(* Logix 5000 project; controller CIP vendor 1 type 14 code 106 rev 20.12; software revision 20.06; part 7 of 13 *)
(* tags used below, declared in another part *)
   Message_Index : ALIAS FOR Integer[30];
   Message_Present : INT[4];
   Message_SEQ : DINT[101];
   Message_Timer : TIMER[1];
   OpCode_Pin : DINT[5];
   PV_Message : DINT[3];
   SCLD_Drain_PH : REAL;
   SCLD_Dryer_Duct_Temp : REAL;
   SCLD_Dryer_Exhaust_Temp : REAL;
   SCLD_Return_Temp : REAL;
   SCLD_Rinse_Cond : REAL;
   SCLD_Solution_Tank_Lvl : REAL;
   SCLD_Solution_Tank_Lvl_Raw : REAL;
   SCLD_Supply_Flow : REAL;
   SCLD_Supply_Flow_CIP : REAL;
   SCLD_Supply_Flow_CIP100 : REAL;
   SCLD_Supply_Flow_CIP200 : REAL;
   SCLD_Supply_Pressure : REAL;
   SCLD_Supply_Temp : REAL;
   SCLD_Wash_Chamber_Lvl : REAL;
   SCLD_Wash_Chamber_Lvl_Raw : REAL;
   SCLD_Wash_Cond : REAL;
   Sequencer : CONTROL[4];
   Solution_Tank_Lvl_Calc : REAL[20];
   Solution_Tank_Lvl_Storage : REAL[3];
   Wash_Chamber_Lvl_Calc : REAL[30];
   Wash_Chamber_Lvl_Storage : REAL[3];
(* MainProgram, continued *)

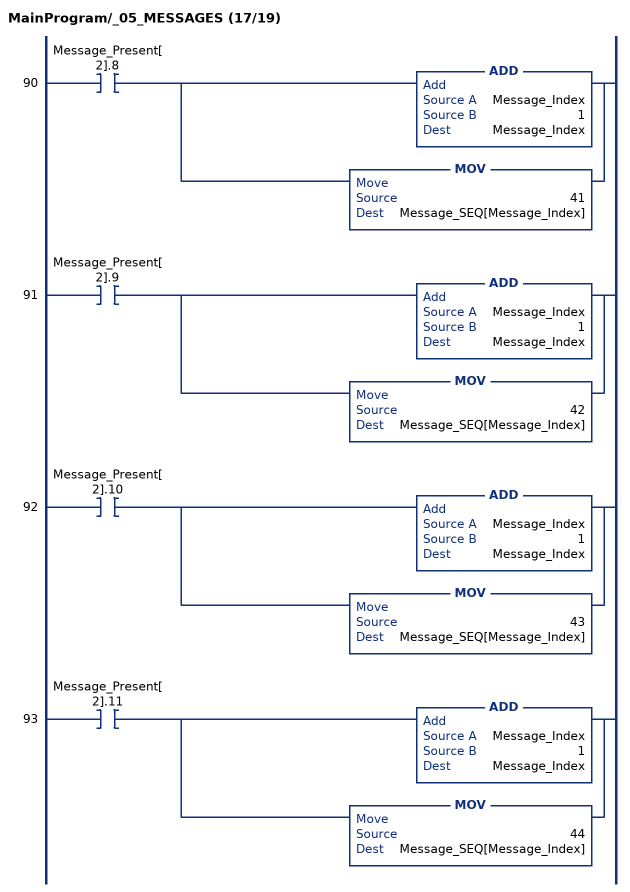
   [picture p115: MainProgram/_05_MESSAGES rungs 90-93]
   90: XIC(Message_Present[2].8)[ADD(Message_Index,1,Message_Index) ,MOV(41,Message_SEQ[Message_Index]) ];
   91: XIC(Message_Present[2].9)[ADD(Message_Index,1,Message_Index) ,MOV(42,Message_SEQ[Message_Index]) ];
   92: XIC(Message_Present[2].10)[ADD(Message_Index,1,Message_Index) ,MOV(43,Message_SEQ[Message_Index]) ];
   93: XIC(Message_Present[2].11)[ADD(Message_Index,1,Message_Index) ,MOV(44,Message_SEQ[Message_Index]) ];
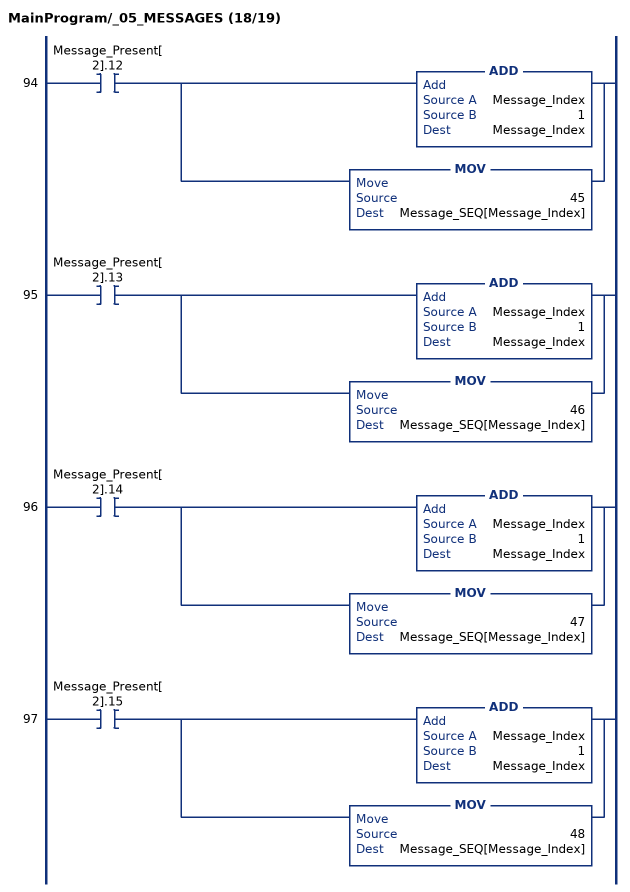
   94: XIC(Message_Present[2].12)[ADD(Message_Index,1,Message_Index) ,MOV(45,Message_SEQ[Message_Index]) ];
   95: XIC(Message_Present[2].13)[ADD(Message_Index,1,Message_Index) ,MOV(46,Message_SEQ[Message_Index]) ];
   96: XIC(Message_Present[2].14)[ADD(Message_Index,1,Message_Index) ,MOV(47,Message_SEQ[Message_Index]) ];
   97: XIC(Message_Present[2].15)[ADD(Message_Index,1,Message_Index) ,MOV(48,Message_SEQ[Message_Index]) ];
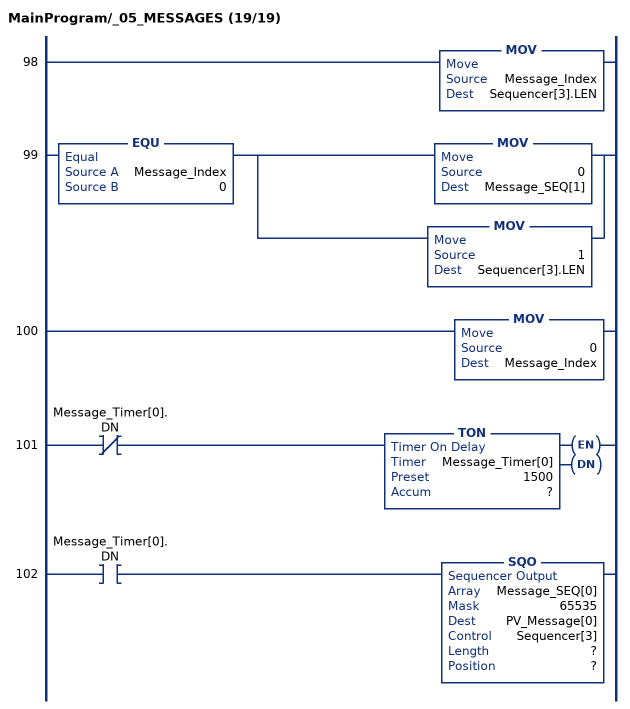
   98: MOV(Message_Index,Sequencer[3].LEN);
   99: EQU(Message_Index,0)[MOV(0,Message_SEQ[1]) ,MOV(1,Sequencer[3].LEN) ];
   100: MOV(0,Message_Index);
   101: XIO(Message_Timer[0].DN)TON(Message_Timer[0],?,?);
   102: XIC(Message_Timer[0].DN)SQO(Message_SEQ[0],65535,PV_Message[0],Sequencer[3],?,?);
END_ROUTINE

ROUTINE _07_SCALE   (* function block diagram *)
   SHEET 1   // Local Analog Input Scaling
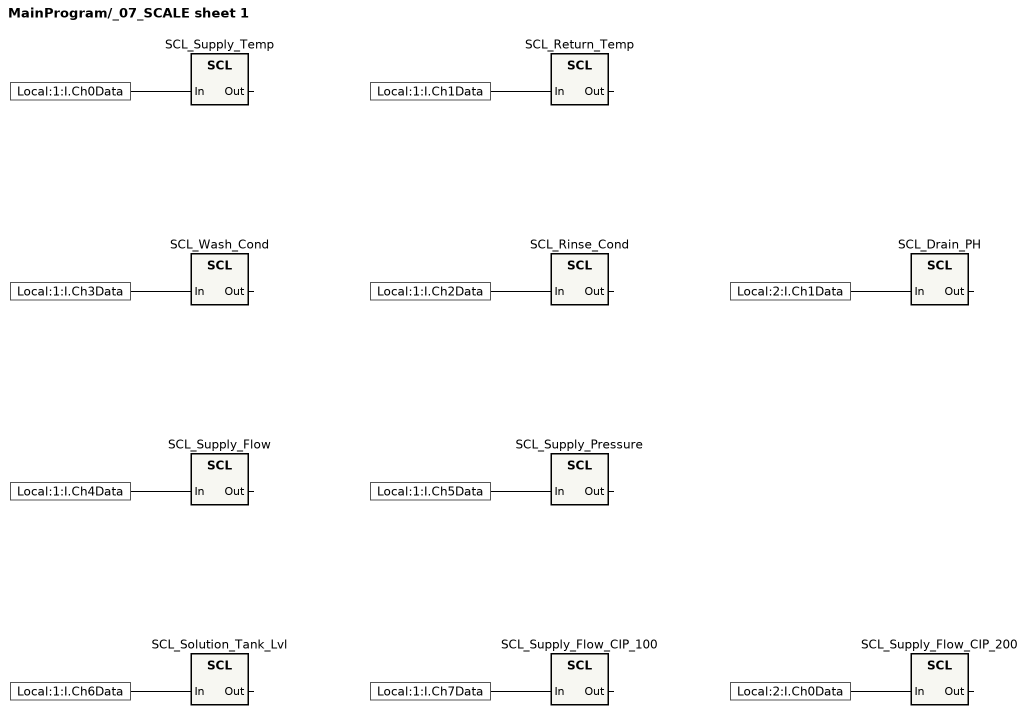
   SCL_Supply_Temp : SCL(In := Local:1:I.Ch0Data);   // unwired pins: Out
   SCL_Wash_Cond : SCL(In := Local:1:I.Ch3Data);   // unwired pins: Out
   SCL_Supply_Flow : SCL(In := Local:1:I.Ch4Data);   // unwired pins: Out
   SCL_Solution_Tank_Lvl : SCL(In := Local:1:I.Ch6Data);   // unwired pins: Out
   SCL_Return_Temp : SCL(In := Local:1:I.Ch1Data);   // unwired pins: Out
   SCL_Rinse_Cond : SCL(In := Local:1:I.Ch2Data);   // unwired pins: Out
   SCL_Supply_Pressure : SCL(In := Local:1:I.Ch5Data);   // unwired pins: Out
   SCL_Supply_Flow_CIP_100 : SCL(In := Local:1:I.Ch7Data);   // unwired pins: Out
   SCL_Drain_PH : SCL(In := Local:2:I.Ch1Data);   // unwired pins: Out
   SCL_Supply_Flow_CIP_200 : SCL(In := Local:2:I.Ch0Data);   // unwired pins: Out
   SHEET 2   // Washer Analog Input Scaling
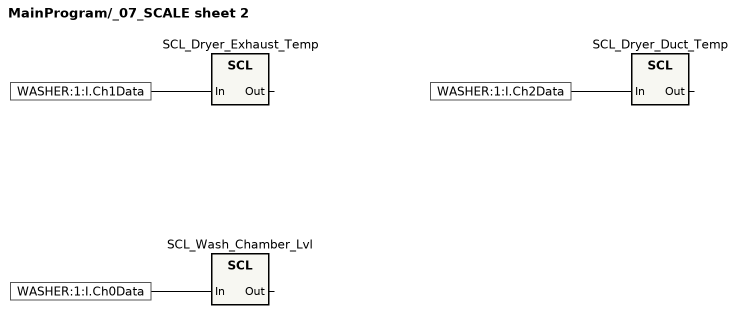
   SCL_Dryer_Exhaust_Temp : SCL(In := WASHER:1:I.Ch1Data);   // unwired pins: Out
   SCL_Wash_Chamber_Lvl : SCL(In := WASHER:1:I.Ch0Data);   // unwired pins: Out
   SCL_Dryer_Duct_Temp : SCL(In := WASHER:1:I.Ch2Data);   // unwired pins: Out
END_ROUTINE

ROUTINE _07_SCALED   (* ladder *)
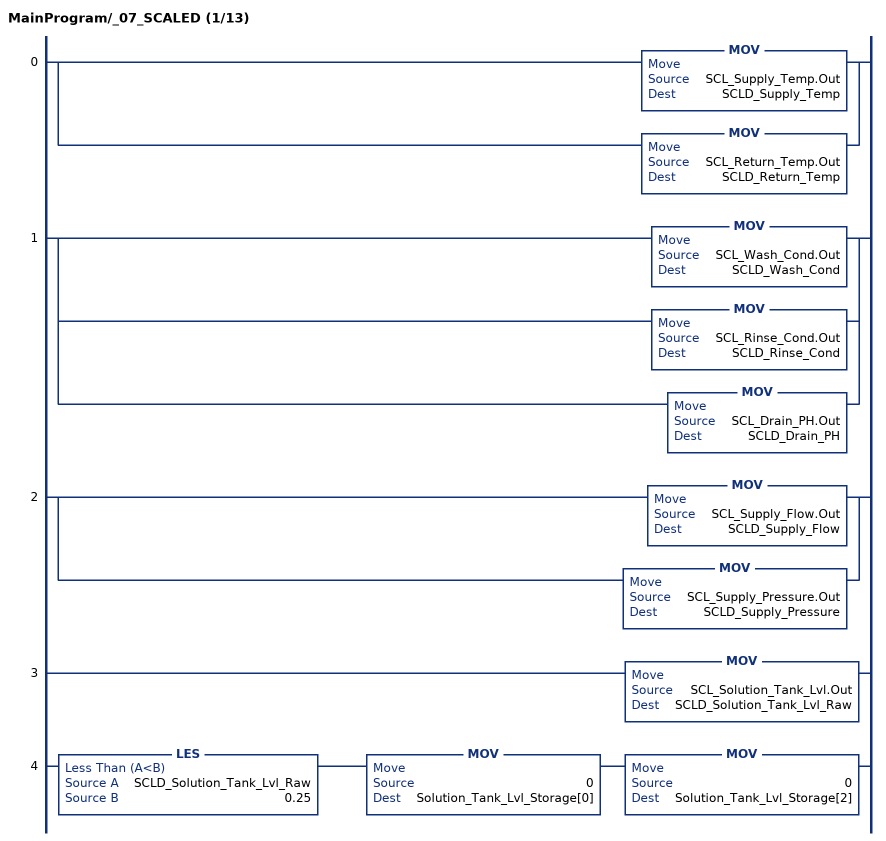
   0: [MOV(SCL_Supply_Temp.Out,SCLD_Supply_Temp) ,MOV(SCL_Return_Temp.Out,SCLD_Return_Temp) ];
   1: [MOV(SCL_Wash_Cond.Out,SCLD_Wash_Cond) ,MOV(SCL_Rinse_Cond.Out,SCLD_Rinse_Cond) ,MOV(SCL_Drain_PH.Out,SCLD_Drain_PH) ];
   2: [MOV(SCL_Supply_Flow.Out,SCLD_Supply_Flow) ,MOV(SCL_Supply_Pressure.Out,SCLD_Supply_Pressure) ];
   3: MOV(SCL_Solution_Tank_Lvl.Out,SCLD_Solution_Tank_Lvl_Raw);
   4: LES(SCLD_Solution_Tank_Lvl_Raw,0.25)MOV(0,Solution_Tank_Lvl_Storage[0])MOV(0,Solution_Tank_Lvl_Storage[2]);
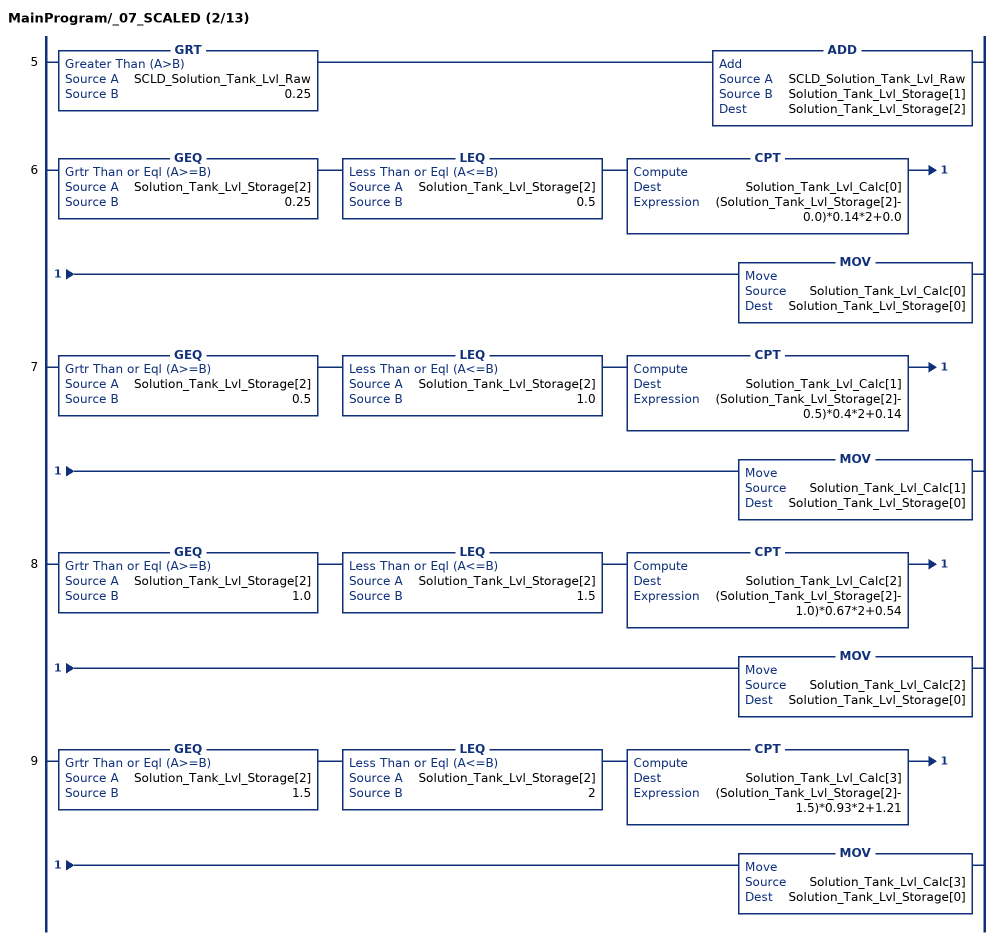
   5: GRT(SCLD_Solution_Tank_Lvl_Raw,0.25)ADD(SCLD_Solution_Tank_Lvl_Raw,Solution_Tank_Lvl_Storage[1],Solution_Tank_Lvl_Storage[2]);
   6: GEQ(Solution_Tank_Lvl_Storage[2],0.25)LEQ(Solution_Tank_Lvl_Storage[2],0.5)CPT(Solution_Tank_Lvl_Calc[0],(Solution_Tank_Lvl_Storage[2]-0.0)*0.14*2+0.0)MOV(Solution_Tank_Lvl_Calc[0],Solution_Tank_Lvl_Storage[0]);
   7: GEQ(Solution_Tank_Lvl_Storage[2],0.5)LEQ(Solution_Tank_Lvl_Storage[2],1.0)CPT(Solution_Tank_Lvl_Calc[1],(Solution_Tank_Lvl_Storage[2]-0.5)*0.4*2+0.14)MOV(Solution_Tank_Lvl_Calc[1],Solution_Tank_Lvl_Storage[0]);
   8: GEQ(Solution_Tank_Lvl_Storage[2],1.0)LEQ(Solution_Tank_Lvl_Storage[2],1.5)CPT(Solution_Tank_Lvl_Calc[2],(Solution_Tank_Lvl_Storage[2]-1.0)*0.67*2+0.54)MOV(Solution_Tank_Lvl_Calc[2],Solution_Tank_Lvl_Storage[0]);
   9: GEQ(Solution_Tank_Lvl_Storage[2],1.5)LEQ(Solution_Tank_Lvl_Storage[2],2)CPT(Solution_Tank_Lvl_Calc[3],(Solution_Tank_Lvl_Storage[2]-1.5)*0.93*2+1.21)MOV(Solution_Tank_Lvl_Calc[3],Solution_Tank_Lvl_Storage[0]);
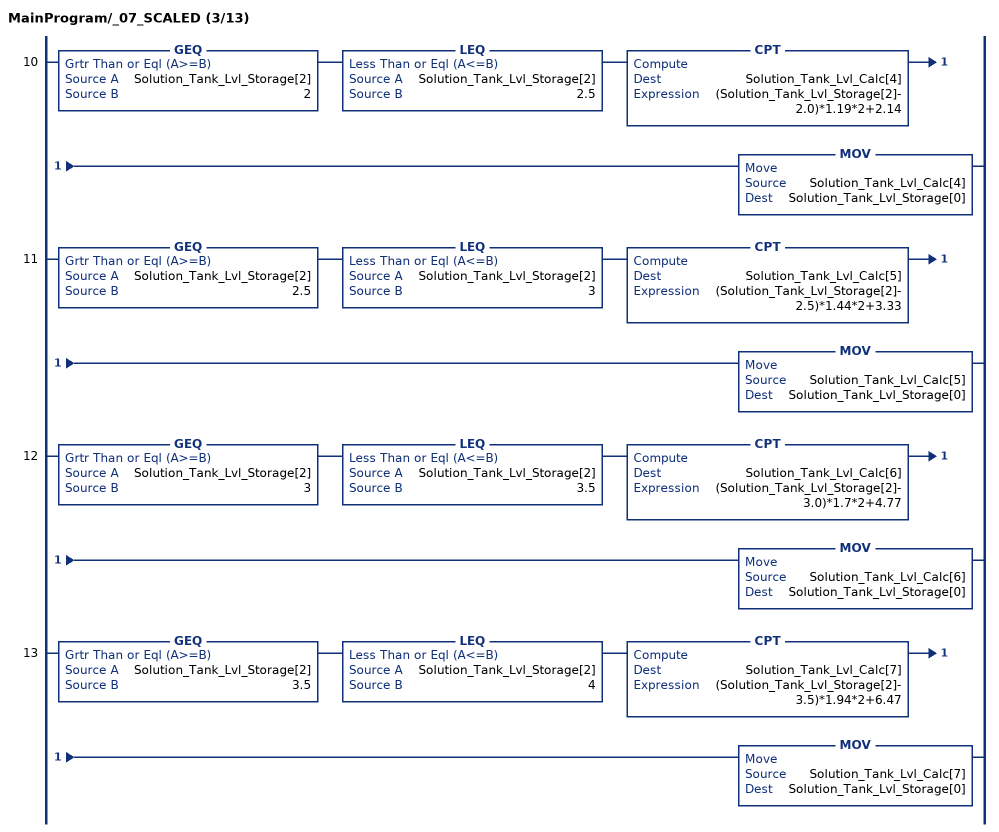
   10: GEQ(Solution_Tank_Lvl_Storage[2],2)LEQ(Solution_Tank_Lvl_Storage[2],2.5)CPT(Solution_Tank_Lvl_Calc[4],(Solution_Tank_Lvl_Storage[2]-2.0)*1.19*2+2.14)MOV(Solution_Tank_Lvl_Calc[4],Solution_Tank_Lvl_Storage[0]);
   11: GEQ(Solution_Tank_Lvl_Storage[2],2.5)LEQ(Solution_Tank_Lvl_Storage[2],3)CPT(Solution_Tank_Lvl_Calc[5],(Solution_Tank_Lvl_Storage[2]-2.5)*1.44*2+3.33)MOV(Solution_Tank_Lvl_Calc[5],Solution_Tank_Lvl_Storage[0]);
   12: GEQ(Solution_Tank_Lvl_Storage[2],3)LEQ(Solution_Tank_Lvl_Storage[2],3.5)CPT(Solution_Tank_Lvl_Calc[6],(Solution_Tank_Lvl_Storage[2]-3.0)*1.7*2+4.77)MOV(Solution_Tank_Lvl_Calc[6],Solution_Tank_Lvl_Storage[0]);
   13: GEQ(Solution_Tank_Lvl_Storage[2],3.5)LEQ(Solution_Tank_Lvl_Storage[2],4)CPT(Solution_Tank_Lvl_Calc[7],(Solution_Tank_Lvl_Storage[2]-3.5)*1.94*2+6.47)MOV(Solution_Tank_Lvl_Calc[7],Solution_Tank_Lvl_Storage[0]);
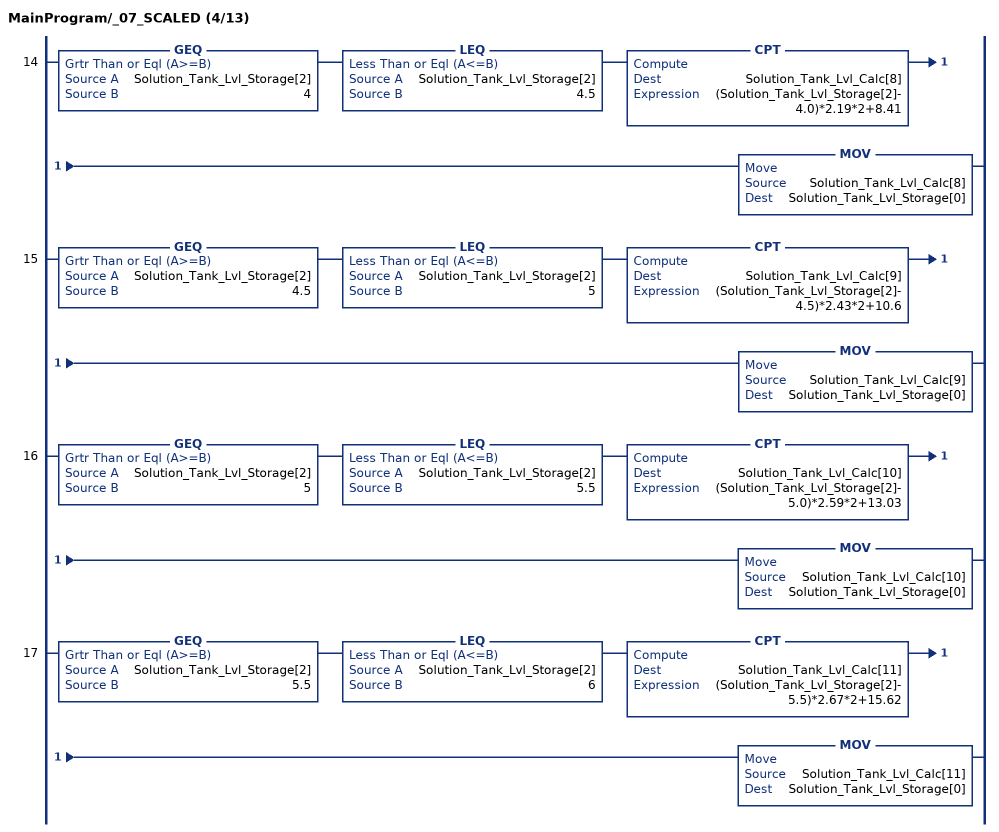
   14: GEQ(Solution_Tank_Lvl_Storage[2],4)LEQ(Solution_Tank_Lvl_Storage[2],4.5)CPT(Solution_Tank_Lvl_Calc[8],(Solution_Tank_Lvl_Storage[2]-4.0)*2.19*2+8.41)MOV(Solution_Tank_Lvl_Calc[8],Solution_Tank_Lvl_Storage[0]);
   15: GEQ(Solution_Tank_Lvl_Storage[2],4.5)LEQ(Solution_Tank_Lvl_Storage[2],5)CPT(Solution_Tank_Lvl_Calc[9],(Solution_Tank_Lvl_Storage[2]-4.5)*2.43*2+10.6)MOV(Solution_Tank_Lvl_Calc[9],Solution_Tank_Lvl_Storage[0]);
   16: GEQ(Solution_Tank_Lvl_Storage[2],5)LEQ(Solution_Tank_Lvl_Storage[2],5.5)CPT(Solution_Tank_Lvl_Calc[10],(Solution_Tank_Lvl_Storage[2]-5.0)*2.59*2+13.03)MOV(Solution_Tank_Lvl_Calc[10],Solution_Tank_Lvl_Storage[0]);
   17: GEQ(Solution_Tank_Lvl_Storage[2],5.5)LEQ(Solution_Tank_Lvl_Storage[2],6)CPT(Solution_Tank_Lvl_Calc[11],(Solution_Tank_Lvl_Storage[2]-5.5)*2.67*2+15.62)MOV(Solution_Tank_Lvl_Calc[11],Solution_Tank_Lvl_Storage[0]);
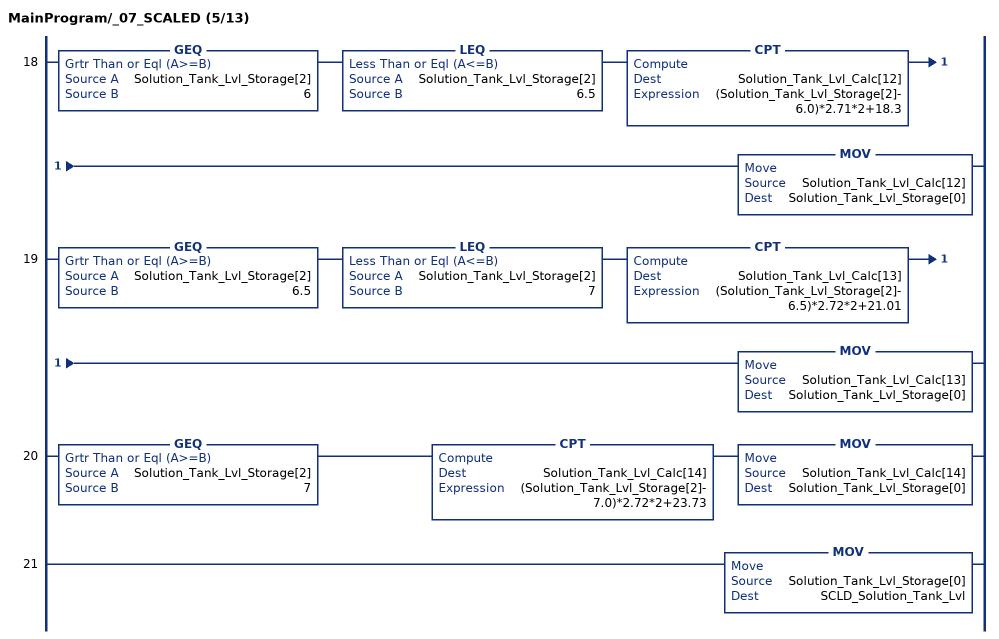
   18: GEQ(Solution_Tank_Lvl_Storage[2],6)LEQ(Solution_Tank_Lvl_Storage[2],6.5)CPT(Solution_Tank_Lvl_Calc[12],(Solution_Tank_Lvl_Storage[2]-6.0)*2.71*2+18.3)MOV(Solution_Tank_Lvl_Calc[12],Solution_Tank_Lvl_Storage[0]);
   19: GEQ(Solution_Tank_Lvl_Storage[2],6.5)LEQ(Solution_Tank_Lvl_Storage[2],7)CPT(Solution_Tank_Lvl_Calc[13],(Solution_Tank_Lvl_Storage[2]-6.5)*2.72*2+21.01)MOV(Solution_Tank_Lvl_Calc[13],Solution_Tank_Lvl_Storage[0]);
   20: GEQ(Solution_Tank_Lvl_Storage[2],7)CPT(Solution_Tank_Lvl_Calc[14],(Solution_Tank_Lvl_Storage[2]-7.0)*2.72*2+23.73)MOV(Solution_Tank_Lvl_Calc[14],Solution_Tank_Lvl_Storage[0]);
   21: MOV(Solution_Tank_Lvl_Storage[0],SCLD_Solution_Tank_Lvl);
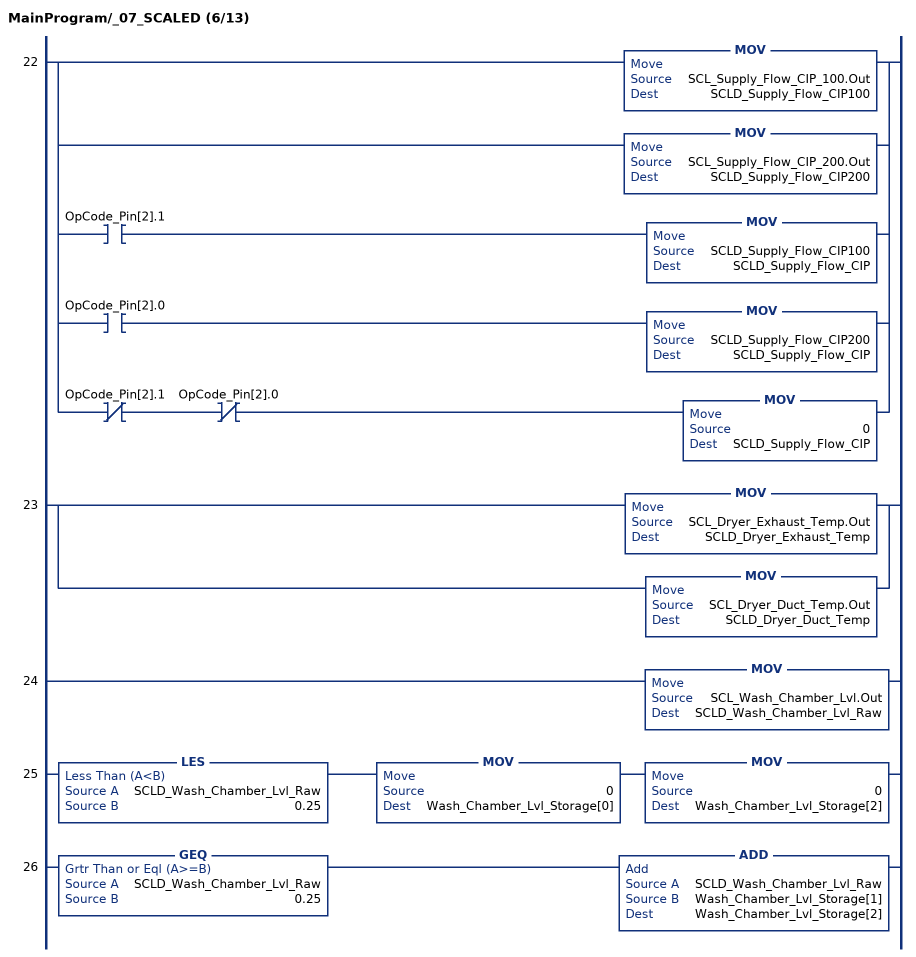
   22: [MOV(SCL_Supply_Flow_CIP_100.Out,SCLD_Supply_Flow_CIP100) ,MOV(SCL_Supply_Flow_CIP_200.Out,SCLD_Supply_Flow_CIP200) ,XIC(OpCode_Pin[2].1) MOV(SCLD_Supply_Flow_CIP100,SCLD_Supply_Flow_CIP) ,XIC(OpCode_Pin[2].0) MOV(SCLD_Supply_Flow_CIP200,SCLD_Supply_Flow_CIP) ,XIO(OpCode_Pin[2].1) XIO(OpCode_Pin[2].0) MOV(0,SCLD_Supply_Flow_CIP) ];
   23: [MOV(SCL_Dryer_Exhaust_Temp.Out,SCLD_Dryer_Exhaust_Temp) ,MOV(SCL_Dryer_Duct_Temp.Out,SCLD_Dryer_Duct_Temp) ];
   24: MOV(SCL_Wash_Chamber_Lvl.Out,SCLD_Wash_Chamber_Lvl_Raw);
   25: LES(SCLD_Wash_Chamber_Lvl_Raw,0.25)MOV(0,Wash_Chamber_Lvl_Storage[0])MOV(0,Wash_Chamber_Lvl_Storage[2]);
   26: GEQ(SCLD_Wash_Chamber_Lvl_Raw,0.25)ADD(SCLD_Wash_Chamber_Lvl_Raw,Wash_Chamber_Lvl_Storage[1],Wash_Chamber_Lvl_Storage[2]);
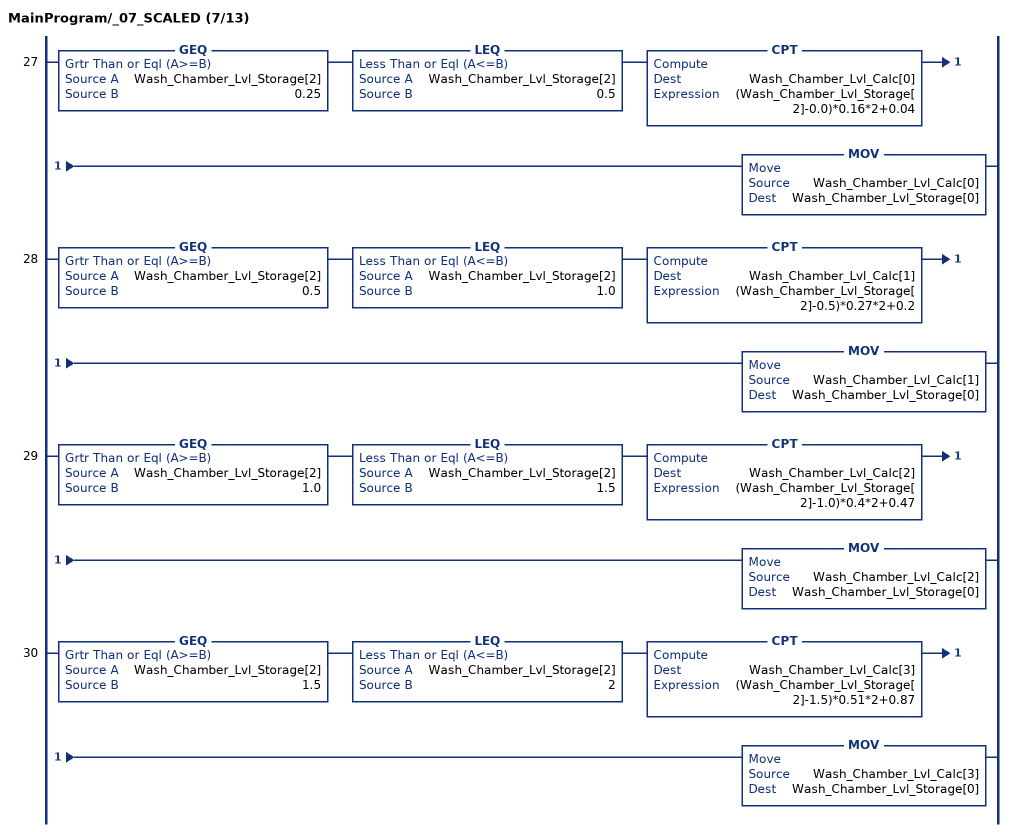
   27: GEQ(Wash_Chamber_Lvl_Storage[2],0.25)LEQ(Wash_Chamber_Lvl_Storage[2],0.5)CPT(Wash_Chamber_Lvl_Calc[0],(Wash_Chamber_Lvl_Storage[2]-0.0)*0.16*2+0.04)MOV(Wash_Chamber_Lvl_Calc[0],Wash_Chamber_Lvl_Storage[0]);
   28: GEQ(Wash_Chamber_Lvl_Storage[2],0.5)LEQ(Wash_Chamber_Lvl_Storage[2],1.0)CPT(Wash_Chamber_Lvl_Calc[1],(Wash_Chamber_Lvl_Storage[2]-0.5)*0.27*2+0.2)MOV(Wash_Chamber_Lvl_Calc[1],Wash_Chamber_Lvl_Storage[0]);
   29: GEQ(Wash_Chamber_Lvl_Storage[2],1.0)LEQ(Wash_Chamber_Lvl_Storage[2],1.5)CPT(Wash_Chamber_Lvl_Calc[2],(Wash_Chamber_Lvl_Storage[2]-1.0)*0.4*2+0.47)MOV(Wash_Chamber_Lvl_Calc[2],Wash_Chamber_Lvl_Storage[0]);
   30: GEQ(Wash_Chamber_Lvl_Storage[2],1.5)LEQ(Wash_Chamber_Lvl_Storage[2],2)CPT(Wash_Chamber_Lvl_Calc[3],(Wash_Chamber_Lvl_Storage[2]-1.5)*0.51*2+0.87)MOV(Wash_Chamber_Lvl_Calc[3],Wash_Chamber_Lvl_Storage[0]);
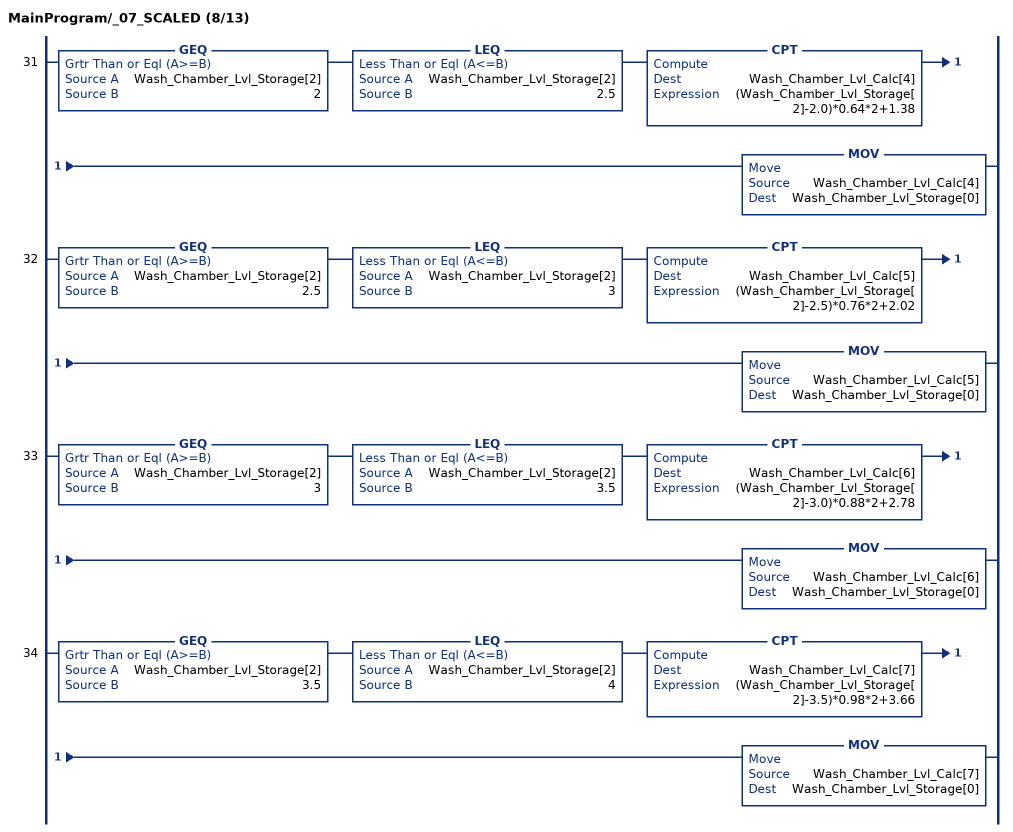
   31: GEQ(Wash_Chamber_Lvl_Storage[2],2)LEQ(Wash_Chamber_Lvl_Storage[2],2.5)CPT(Wash_Chamber_Lvl_Calc[4],(Wash_Chamber_Lvl_Storage[2]-2.0)*0.64*2+1.38)MOV(Wash_Chamber_Lvl_Calc[4],Wash_Chamber_Lvl_Storage[0]);
   32: GEQ(Wash_Chamber_Lvl_Storage[2],2.5)LEQ(Wash_Chamber_Lvl_Storage[2],3)CPT(Wash_Chamber_Lvl_Calc[5],(Wash_Chamber_Lvl_Storage[2]-2.5)*0.76*2+2.02)MOV(Wash_Chamber_Lvl_Calc[5],Wash_Chamber_Lvl_Storage[0]);
   33: GEQ(Wash_Chamber_Lvl_Storage[2],3)LEQ(Wash_Chamber_Lvl_Storage[2],3.5)CPT(Wash_Chamber_Lvl_Calc[6],(Wash_Chamber_Lvl_Storage[2]-3.0)*0.88*2+2.78)MOV(Wash_Chamber_Lvl_Calc[6],Wash_Chamber_Lvl_Storage[0]);
   34: GEQ(Wash_Chamber_Lvl_Storage[2],3.5)LEQ(Wash_Chamber_Lvl_Storage[2],4)CPT(Wash_Chamber_Lvl_Calc[7],(Wash_Chamber_Lvl_Storage[2]-3.5)*0.98*2+3.66)MOV(Wash_Chamber_Lvl_Calc[7],Wash_Chamber_Lvl_Storage[0]);
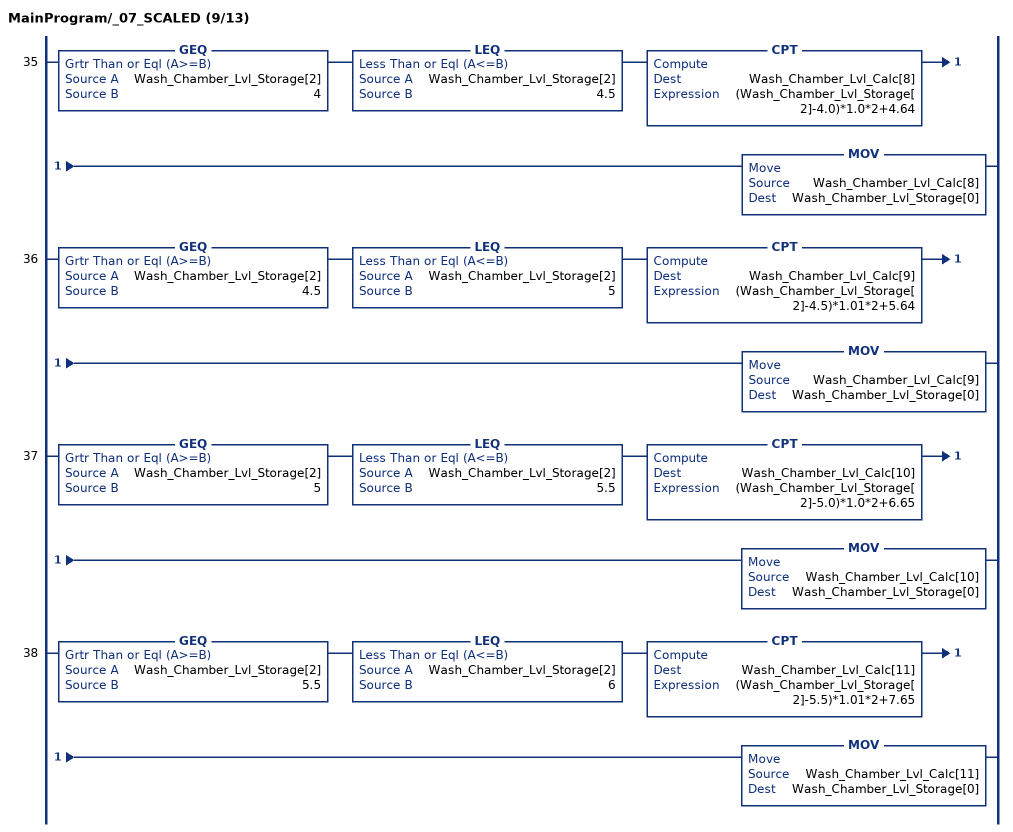
   35: GEQ(Wash_Chamber_Lvl_Storage[2],4)LEQ(Wash_Chamber_Lvl_Storage[2],4.5)CPT(Wash_Chamber_Lvl_Calc[8],(Wash_Chamber_Lvl_Storage[2]-4.0)*1.0*2+4.64)MOV(Wash_Chamber_Lvl_Calc[8],Wash_Chamber_Lvl_Storage[0]);
   36: GEQ(Wash_Chamber_Lvl_Storage[2],4.5)LEQ(Wash_Chamber_Lvl_Storage[2],5)CPT(Wash_Chamber_Lvl_Calc[9],(Wash_Chamber_Lvl_Storage[2]-4.5)*1.01*2+5.64)MOV(Wash_Chamber_Lvl_Calc[9],Wash_Chamber_Lvl_Storage[0]);
   37: GEQ(Wash_Chamber_Lvl_Storage[2],5)LEQ(Wash_Chamber_Lvl_Storage[2],5.5)CPT(Wash_Chamber_Lvl_Calc[10],(Wash_Chamber_Lvl_Storage[2]-5.0)*1.0*2+6.65)MOV(Wash_Chamber_Lvl_Calc[10],Wash_Chamber_Lvl_Storage[0]);
   38: GEQ(Wash_Chamber_Lvl_Storage[2],5.5)LEQ(Wash_Chamber_Lvl_Storage[2],6)CPT(Wash_Chamber_Lvl_Calc[11],(Wash_Chamber_Lvl_Storage[2]-5.5)*1.01*2+7.65)MOV(Wash_Chamber_Lvl_Calc[11],Wash_Chamber_Lvl_Storage[0]);
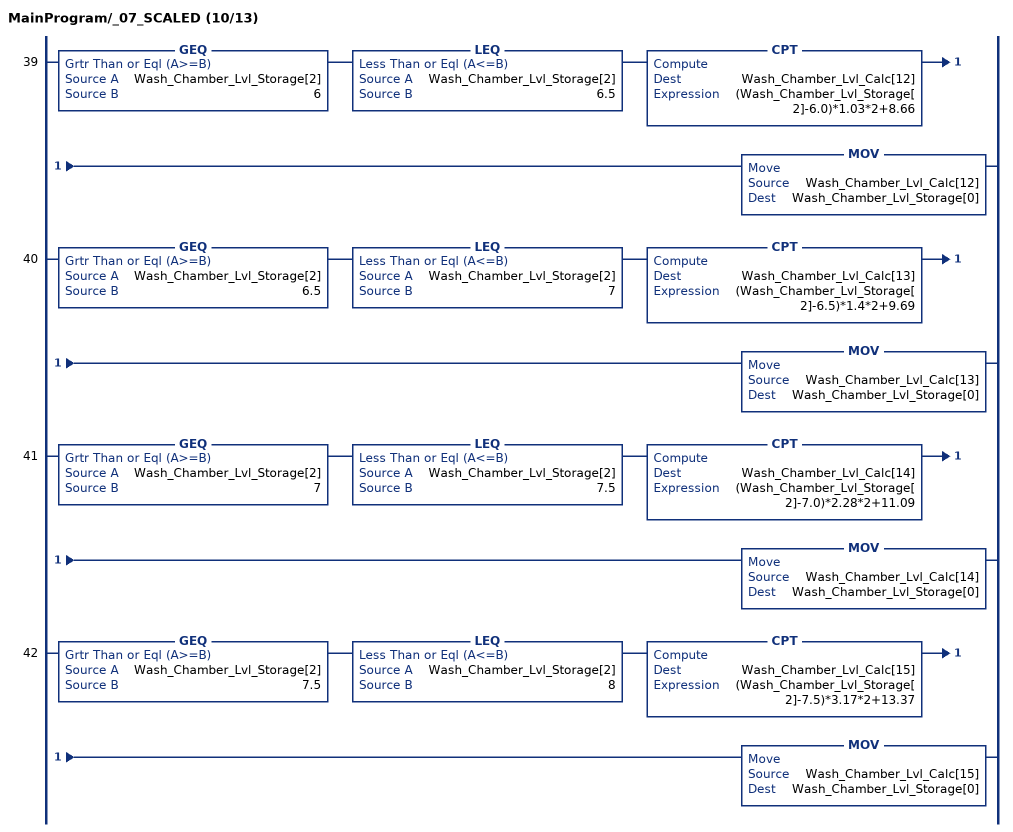
   39: GEQ(Wash_Chamber_Lvl_Storage[2],6)LEQ(Wash_Chamber_Lvl_Storage[2],6.5)CPT(Wash_Chamber_Lvl_Calc[12],(Wash_Chamber_Lvl_Storage[2]-6.0)*1.03*2+8.66)MOV(Wash_Chamber_Lvl_Calc[12],Wash_Chamber_Lvl_Storage[0]);
   40: GEQ(Wash_Chamber_Lvl_Storage[2],6.5)LEQ(Wash_Chamber_Lvl_Storage[2],7)CPT(Wash_Chamber_Lvl_Calc[13],(Wash_Chamber_Lvl_Storage[2]-6.5)*1.4*2+9.69)MOV(Wash_Chamber_Lvl_Calc[13],Wash_Chamber_Lvl_Storage[0]);
   41: GEQ(Wash_Chamber_Lvl_Storage[2],7)LEQ(Wash_Chamber_Lvl_Storage[2],7.5)CPT(Wash_Chamber_Lvl_Calc[14],(Wash_Chamber_Lvl_Storage[2]-7.0)*2.28*2+11.09)MOV(Wash_Chamber_Lvl_Calc[14],Wash_Chamber_Lvl_Storage[0]);
   42: GEQ(Wash_Chamber_Lvl_Storage[2],7.5)LEQ(Wash_Chamber_Lvl_Storage[2],8)CPT(Wash_Chamber_Lvl_Calc[15],(Wash_Chamber_Lvl_Storage[2]-7.5)*3.17*2+13.37)MOV(Wash_Chamber_Lvl_Calc[15],Wash_Chamber_Lvl_Storage[0]);
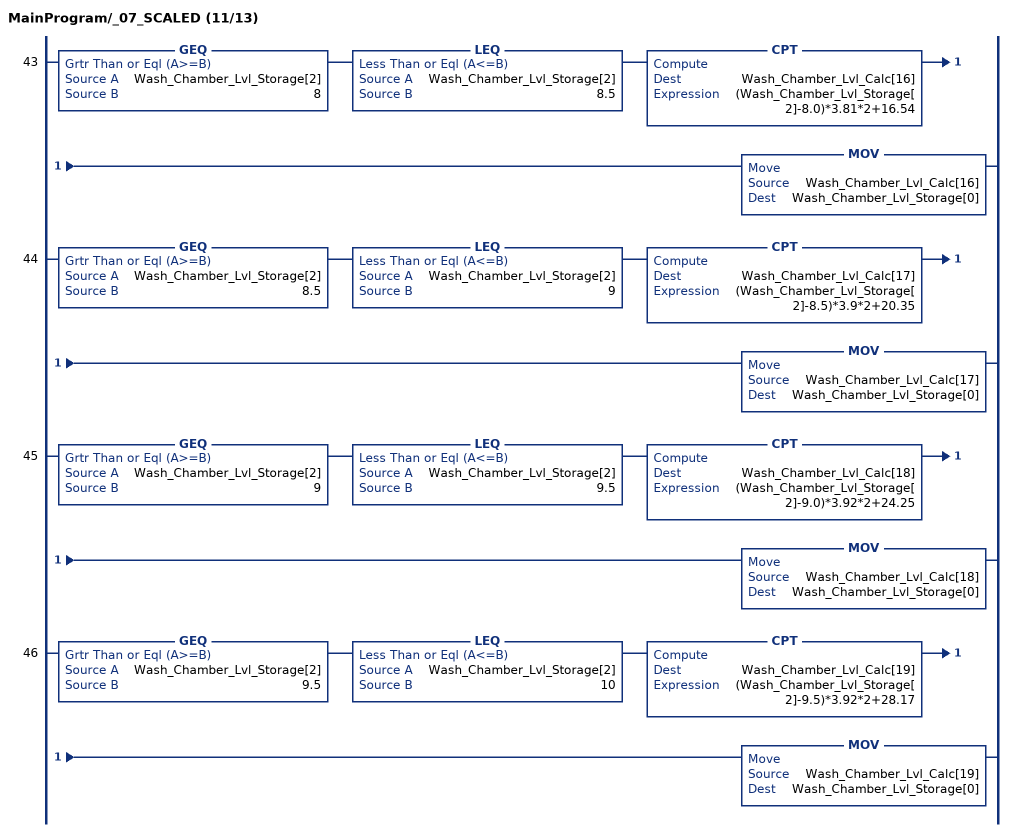
   43: GEQ(Wash_Chamber_Lvl_Storage[2],8)LEQ(Wash_Chamber_Lvl_Storage[2],8.5)CPT(Wash_Chamber_Lvl_Calc[16],(Wash_Chamber_Lvl_Storage[2]-8.0)*3.81*2+16.54)MOV(Wash_Chamber_Lvl_Calc[16],Wash_Chamber_Lvl_Storage[0]);
   44: GEQ(Wash_Chamber_Lvl_Storage[2],8.5)LEQ(Wash_Chamber_Lvl_Storage[2],9)CPT(Wash_Chamber_Lvl_Calc[17],(Wash_Chamber_Lvl_Storage[2]-8.5)*3.9*2+20.35)MOV(Wash_Chamber_Lvl_Calc[17],Wash_Chamber_Lvl_Storage[0]);
   45: GEQ(Wash_Chamber_Lvl_Storage[2],9)LEQ(Wash_Chamber_Lvl_Storage[2],9.5)CPT(Wash_Chamber_Lvl_Calc[18],(Wash_Chamber_Lvl_Storage[2]-9.0)*3.92*2+24.25)MOV(Wash_Chamber_Lvl_Calc[18],Wash_Chamber_Lvl_Storage[0]);
   46: GEQ(Wash_Chamber_Lvl_Storage[2],9.5)LEQ(Wash_Chamber_Lvl_Storage[2],10)CPT(Wash_Chamber_Lvl_Calc[19],(Wash_Chamber_Lvl_Storage[2]-9.5)*3.92*2+28.17)MOV(Wash_Chamber_Lvl_Calc[19],Wash_Chamber_Lvl_Storage[0]);
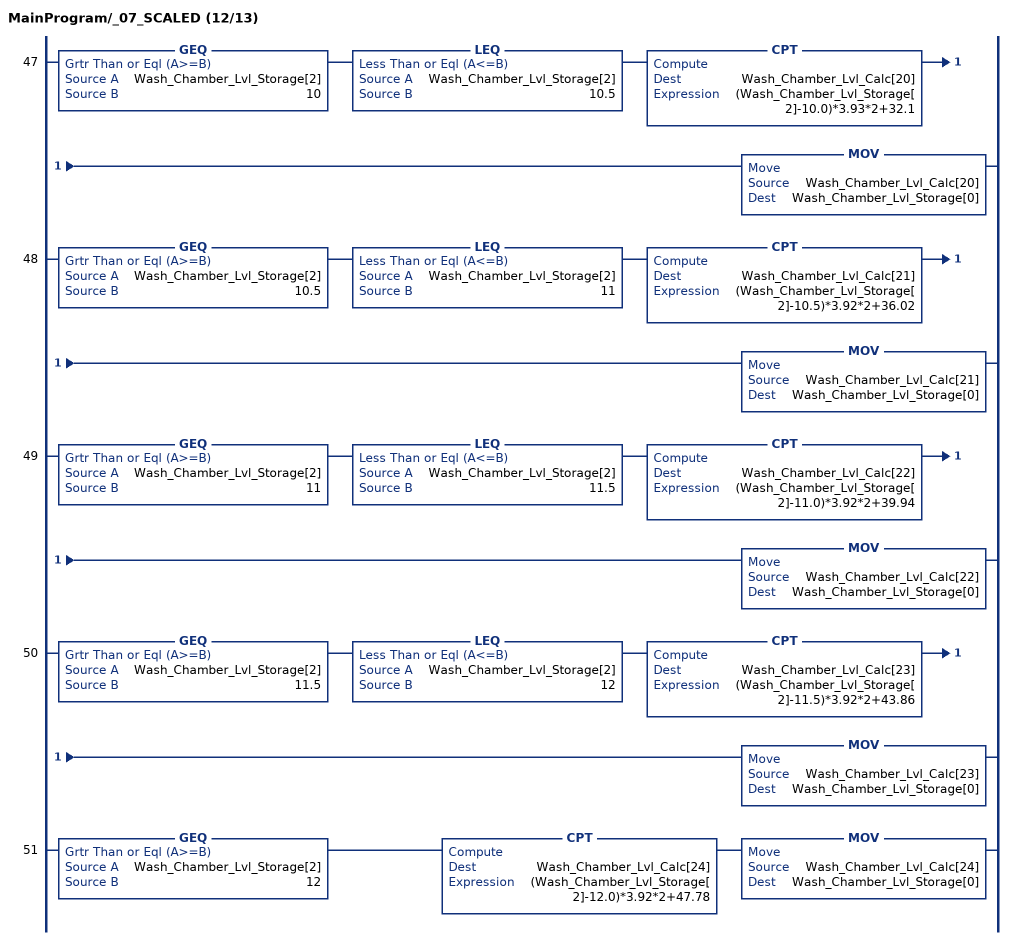
   47: GEQ(Wash_Chamber_Lvl_Storage[2],10)LEQ(Wash_Chamber_Lvl_Storage[2],10.5)CPT(Wash_Chamber_Lvl_Calc[20],(Wash_Chamber_Lvl_Storage[2]-10.0)*3.93*2+32.1)MOV(Wash_Chamber_Lvl_Calc[20],Wash_Chamber_Lvl_Storage[0]);
   48: GEQ(Wash_Chamber_Lvl_Storage[2],10.5)LEQ(Wash_Chamber_Lvl_Storage[2],11)CPT(Wash_Chamber_Lvl_Calc[21],(Wash_Chamber_Lvl_Storage[2]-10.5)*3.92*2+36.02)MOV(Wash_Chamber_Lvl_Calc[21],Wash_Chamber_Lvl_Storage[0]);
   49: GEQ(Wash_Chamber_Lvl_Storage[2],11)LEQ(Wash_Chamber_Lvl_Storage[2],11.5)CPT(Wash_Chamber_Lvl_Calc[22],(Wash_Chamber_Lvl_Storage[2]-11.0)*3.92*2+39.94)MOV(Wash_Chamber_Lvl_Calc[22],Wash_Chamber_Lvl_Storage[0]);
   50: GEQ(Wash_Chamber_Lvl_Storage[2],11.5)LEQ(Wash_Chamber_Lvl_Storage[2],12)CPT(Wash_Chamber_Lvl_Calc[23],(Wash_Chamber_Lvl_Storage[2]-11.5)*3.92*2+43.86)MOV(Wash_Chamber_Lvl_Calc[23],Wash_Chamber_Lvl_Storage[0]);
   51: GEQ(Wash_Chamber_Lvl_Storage[2],12)CPT(Wash_Chamber_Lvl_Calc[24],(Wash_Chamber_Lvl_Storage[2]-12.0)*3.92*2+47.78)MOV(Wash_Chamber_Lvl_Calc[24],Wash_Chamber_Lvl_Storage[0]);
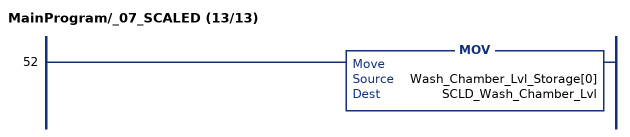
   52: MOV(Wash_Chamber_Lvl_Storage[0],SCLD_Wash_Chamber_Lvl);
END_ROUTINE
